// TIA Portal V21 export
// export: Created 2026-10-12T11:32:17.0003968Z, ExportSetting WithDefaults, DisplayName Totally Integrated Automation Portal, DisplayVersion V21, DisplayName STEP 7 Professional, DisplayVersion V21, DisplayName STEP 7 Safety, DisplayVersion V21, DisplayName Tech WebApplication, DisplayVersion V21, DisplayName WinCC Basic/Comfort/Advanced, DisplayVersion V21, DisplayName WinCC Unified, DisplayVersion V21
DATA_BLOCK "DB_CAMERA"   // DB5
{ S7_Optimized_Access := 'FALSE' }
VERSION : 0.1
// stored: AutoNumber true, DBAccessibleFromOPCUA true, IsOnlyStoredInLoadMemory false, IsWriteProtectedInAS false
   VAR
      DATA1 : Int;
      DATA2 : Int;
      DATA3 : Int;
      DATA4 : Int;
      DATA5 : Int;
      DATA6 : Int;
      DATA7 : Int;
      DATA8 : Int;
      DATA9 : Int;
      DATA10 : Int;
      DATA11 : Int;
      DATA12 : Int;
      DATA13 : Int;
      DATA14 : Int;
      DATA15 : Int;
      DATA16 : Int;
      DATA17 : Int;
      DATA18 : Int;
      DATA19 : Int;
   END_VAR
BEGIN
END_DATA_BLOCK
